(* IEC 61131-3 sources: kns-port-domestic/tools/port_metrics_tests/fixtures/adapted/src/GVLs, 1 file *)

(* ---- GVL_Cfg.gvl.st ---- *)
// PORT: [io] конфигурация насосов для каналов REGUL
// PORT: [hmi]
{attribute 'qualified_only'}
VAR_GLOBAL
    stPump : ST_PumpCfg;
END_VAR
